// TIA Portal project "Test_PID_Compact_Factory_Cuve" (V16)

(* hardware
DEVICE "Station S7-1200_1"  S7-1200 Station
   slot 0: "Châssis_0"  S7-1200 Rack  Rack  V1.0
   slot 1: "PLC_1"  CPU 1212C DC/DC/DC  6ES7 212-1AE40-0XB0  V4.4
DEVICE "HMI_1"  KTP1200 Basic PN
   slot 0: "HMI_1"  KTP1200 Basic PN  6AV2 123-2MB03-0AX0  16.0.0.0
   slot 1: "HMI_RT_1"  KTP1200 Basic PN  6AV2 123-2MB03-0AX0  16.0.0.0
   slot 5: "HMI_1.IE_CP_1"  PROFINET Interface  16.0.0.0
      slot 1: "Interface PROFINET_1"  PROFINET Interface
         slot 1: "Port_1"  Port
*)

// ===== PLC "PLC_1"  CPU 1212C DC/DC/DC =====

VAR_GLOBAL   // PLC tag table "Table de variables standard"
   "Clock_Byte" AT %MB1000 : Byte;
   "Clock_10Hz" AT %M1000.0 : Bool;
   "Clock_5Hz" AT %M1000.1 : Bool;
   "Clock_2.5Hz" AT %M1000.2 : Bool;
   "Clock_2Hz" AT %M1000.3 : Bool;
   "Clock_1.25Hz" AT %M1000.4 : Bool;
   "Clock_1Hz" AT %M1000.5 : Bool;
   "Clock_0.625Hz" AT %M1000.6 : Bool;
   "Clock_0.5Hz" AT %M1000.7 : Bool;
   "Bouton_0" AT %I0.0 : Bool;
   "Bouton_1" AT %I0.1 : Bool;
   "Bouton_2" AT %I0.2 : Bool;
   "Bouton_3" AT %I0.3 : Bool;
   "Bouton_4" AT %I0.4 : Bool;
   "Bouton_5" AT %I0.5 : Bool;
   "Bouton_6" AT %I0.6 : Bool;
   "Bouton_7" AT %I0.7 : Bool;
   "Sortie_0" AT %Q0.0 : Bool;
   "Sortie_1" AT %Q0.1 : Bool;
   "Sortie_2" AT %Q0.2 : Bool;
   "Sortie_3" AT %Q0.3 : Bool;
   "Sortie_4" AT %Q0.4 : Bool;
   "Sortie_5" AT %Q0.5 : Bool;
   "Commande_Vanne_pcent" AT %MD6 : Real;
   "Consigne_Niveau_Litres" AT %MD10 : Real;
   "Bruit" AT %MD18 : Real;
   "Erreur_Niveau_Litres" AT %MD22 : Real;
   "Correcteur_P_Coeff" AT %MD30 : Real;
   "Erreur_Niveau_pcent" AT %MD26 : Real;
   "Limite_Commande_Max_pcent" AT %MD34 : Real;
   "Limite_Commande_Min_pcent" AT %MD38 : Real;
   "Commande_Max_Atteinte" AT %M70.0 : Bool;
   "Commande_Min_Atteinte" AT %M70.1 : Bool;
   "Consigne_Niveau_Auto_Max" AT %MD42 : Real;
   "Consigne_Niveau_Auto_Min" AT %MD46 : Real;
   "Duree_Demi_Cycle" AT %MD50 : Time;
   "Duree_Demi_Cycle_sec" AT %MW54 : Int;
   "Correcteur_Ti_Valeur_sec" AT %MD72 : Real;
   "Correcteur_Td_Valeur_sec" AT %MD76 : Real;
   "Correcteur_KP_pondere" AT %MD80 : Real;
   "Correcteur_Td_pondere" AT %MD84 : Real;
   "Correcteur_Fo_PB_Derive" AT %MD88 : Real;
   "Commande_Evacuation_pcent" AT %MD14 : Real;
   "Niveau_Litres" AT %MD92 : Real;
   "Debit_Entree_lpars" AT %MD200 : Real;
   "Debit_Sortie_lpars" AT %MD204 : Real;
   "Correcteur_Coeff_Disturbance" AT %MD208 : Real;
END_VAR

VAR_GLOBAL   // PLC tag table "Table de variables IHM"
   "IHM_Bouton_Oscillo_1" AT %M100.0 : Bool;
   "IHM_Bouton_Oscillo_2" AT %M100.1 : Bool;
   "IHM_Bouton_PID_ON_OFF" AT %M100.2 : Bool;
   "IHM_Bouton_Limit_ON_OFF" AT %M100.3 : Bool;
   "IHM_Bouton_Boucle_Fermee" AT %M100.4 : Bool;
   "IHM_Bouton_Bruit" AT %M100.5 : Bool;
   "IHM_Affichage_Oscillo_2" AT %M112.0 : Bool;
   "IHM_Bouton_Marche_Auto" AT %M100.6 : Bool;
   "IHM_Affichage_Correcteur" AT %M112.1 : Bool;
   "IHM_Affichage_Correcteur_I" AT %M112.4 : Bool;
   "IHM_Affichage_Correcteur_D" AT %M112.5 : Bool;
   "IHM_Bouton_Correcteur_I" AT %M112.2 : Bool;
   "IHM_Bouton_Correcteur_D" AT %M112.3 : Bool;
   "IHM_Curseur_Correcteur_I" AT %M112.6 : Bool;
   "IHM_Curseur_Correcteur_D" AT %M112.7 : Bool;
   "IHM_Curseur_Correcteur_P" AT %M113.1 : Bool;
   "IHM_Affichage_Tuyau_Arrivee" AT %M113.2 : Bool;
   "IHM_Affichage_Tuyau_Evacuation" AT %M113.3 : Bool;
   "IHM_Deplacement_Fleche_Tuyau_Arrivee" AT %MW114 : Int;
   "IHM_Deplacement_Fleche_Tuyau_Evacuation" AT %MW116 : Int;
   "IHM_Bouton_Disturbance" AT %M113.4 : Bool;
   "IHM_Affichage_Correcteur_A" AT %M113.5 : Bool;
   "IHM_Valeur_Disturbance" AT %MD120 : Real;
END_VAR

VAR_GLOBAL   // PLC tag table "Table de variables Factory"
   "Niveau_Cuve_Factory" AT %IW100 : Int;
   "Commande_Vanne_Factory" AT %QW100 : Int;
   "Commande_Evacuation_Factory" AT %QW102 : Int;
   "Debit_Sortie_Factory" AT %IW102 : Int;
   "Warning_Light" AT %Q200.0 : Bool;
END_VAR

// folder: Régulateur

DATA_BLOCK "Regulation_DB"   // DB2
{ S7_Optimized_Access := 'TRUE' }
VERSION : 0.1
// stored: InstanceOfName Regulation
"Regulation"
BEGIN
END_DATA_BLOCK

// folder: Simulation Systeme

DATA_BLOCK "POV_DB"   // DB1
{ S7_Optimized_Access := 'TRUE' }
VERSION : 0.1
// stored: InstanceOfName POV
"POV"
BEGIN
END_DATA_BLOCK

// folder: Régulateur

FUNCTION_BLOCK "Regulation"   // FB2, LAD
{ S7_Optimized_Access := 'TRUE' }
VERSION : 0.1
   VAR_TEMP
      Commande_Anticipatrice : Real;
   END_VAR
BEGIN

REGION Network 1 (SCL): Commande Anticipatrice
   IF "IHM_Bouton_Disturbance" THEN
       IF "Erreur_Niveau_Litres">=-1.0 THEN
           #Commande_Anticipatrice := "Debit_Sortie_lpars" * "Correcteur_Coeff_Disturbance";
       ELSE
           #Commande_Anticipatrice := 0;
       END_IF;
   ELSE
       #Commande_Anticipatrice := 0;
   END_IF;

   "IHM_Valeur_Disturbance" := #Commande_Anticipatrice;
END_REGION

REGION Network 2: Bloc fonction PID_Compact
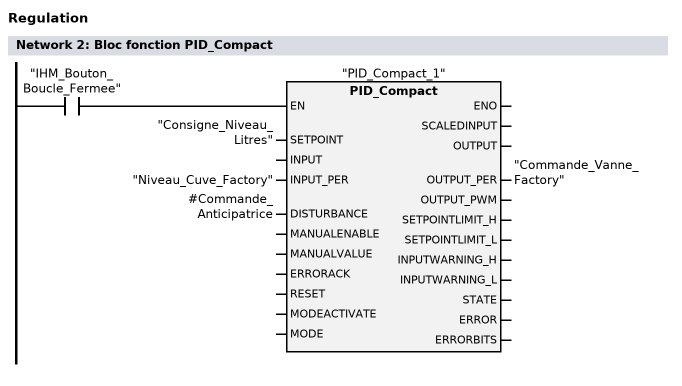
   IF "IHM_Bouton_Boucle_Fermee" THEN
       "PID_Compact_1"(Setpoint := "Consigne_Niveau_Litres",   // PID_Compact
                       Input_PER := "Niveau_Cuve_Factory",
                       Disturbance := #Commande_Anticipatrice,
                       Output_PER => "Commande_Vanne_Factory");
   END_IF;
END_REGION

REGION Network 3 (SCL): Affectation grandeur de commande BO/BF
   // ==== Commande BO / BF ==============================================================================================================
   IF "IHM_Bouton_Boucle_Fermee" THEN
       "Commande_Vanne_pcent":=(INT_TO_REAL("Commande_Vanne_Factory")/27648.0)*100.0;
       "Niveau_Litres" := "PID_Compact_1".ScaledInput;
   ELSE
       "Commande_Vanne_pcent" := "Consigne_Niveau_Litres" ; // Pas des vrais litres...
       "Commande_Vanne_Factory" := REAL_TO_INT("Commande_Vanne_pcent" * 27648.0 / 100.0);
       "Erreur_Niveau_Litres" := 0.0;
       "Erreur_Niveau_pcent" := 0.0;
       "Niveau_Litres" := 300.0 * INT_TO_REAL("Niveau_Cuve_Factory") / 27648.0;
   END_IF;



   // ==== Gestion des limitations de commande ============================================================================================
   REGION Limitations_Commande
       IF "Commande_Vanne_pcent">= "Limite_Commande_Max_pcent" THEN
           "Commande_Vanne_pcent" := "Limite_Commande_Max_pcent";
           "Commande_Max_Atteinte" := "IHM_Bouton_Limit_ON_OFF";
       ELSE
           "Commande_Max_Atteinte" := FALSE;
       END_IF;
       IF "Commande_Vanne_pcent" <= "Limite_Commande_Min_pcent" THEN
           "Commande_Vanne_pcent" := "Limite_Commande_Min_pcent";
           "Commande_Min_Atteinte" := "IHM_Bouton_Limit_ON_OFF";
       ELSE
           "Commande_Min_Atteinte" := FALSE;
       END_IF;
   END_REGION
END_REGION

REGION Network 4 (SCL): Pour affichage IHM
   // ---- Calcul Erreur
   "Erreur_Niveau_Litres" := "Consigne_Niveau_Litres" - "PID_Compact_1".ScaledInput ;
   IF "Consigne_Niveau_Litres" <> 0.0 THEN
       "Erreur_Niveau_pcent" := ("Erreur_Niveau_Litres" / "Consigne_Niveau_Litres") * 100.0;
   ELSE
       "Erreur_Niveau_pcent" := 0.0;
   END_IF;
END_REGION
END_FUNCTION_BLOCK

ORGANIZATION_BLOCK "Appel_Regulation"   // OB32, LAD, CyclicInterrupt
{ S7_Optimized_Access := 'TRUE' }
VERSION : 0.1
   VAR_INPUT
      Initial_Call : Bool;   // Initial call of this OB
      Event_Count : Int;   // Events discarded
   END_VAR
BEGIN

REGION Network 1
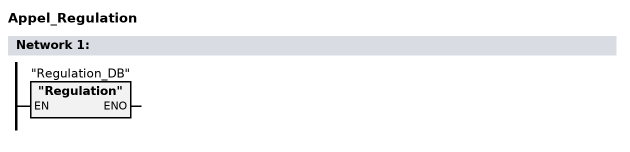
   RUNG wire#powerrail
      "Regulation_DB"()
   END_RUNG
   // the same network as SCL:
   "Regulation_DB"();   // "Regulation"
END_REGION
END_ORGANIZATION_BLOCK

// folder: Simulation Systeme

FUNCTION_BLOCK "POV"   // FB1, LAD
{ S7_Optimized_Access := 'TRUE' }
VERSION : 0.1
   VAR
      Coeff_Perte_Vitesse : Real := 0.3;   // Si 0,4 Perte de 40%
      Temps_Cycle : TON_TIME;
      Temps_Cycle_Demi : TP_TIME;
      Pulse_Cycle : Bool;
   END_VAR
   VAR_TEMP
      Duree_Cycle : Time;
   END_VAR
BEGIN

REGION Network 1 (SCL)
   // ===== Limitations saisie utilisateur IHM =================================================================================

   REGION Limitations_Saisies
       IF "IHM_Bouton_Boucle_Fermee" THEN
           IF "Consigne_Niveau_Litres" > 300.0 THEN
               "Consigne_Niveau_Litres" := 300.0;  // Des vrais litres
           END_IF;
       ELSE
           IF "Consigne_Niveau_Litres" > 100.0 THEN
               "Consigne_Niveau_Litres" := 100.0;  // Pas des litres, mais un pourcentage d'ouverture de la vanne
           END_IF;
           ;
       END_IF;

       IF "Consigne_Niveau_Litres" < 0 THEN
           "Consigne_Niveau_Litres" := 0.0;
       END_IF;

       IF "Commande_Evacuation_pcent" > 100.0 THEN
           "Commande_Evacuation_pcent" := 100.0;
       END_IF;
       IF "Commande_Evacuation_pcent" <0  THEN
           "Commande_Evacuation_pcent" := 0.0;
       END_IF;
   END_REGION


   // ===== Evacuation et débits E/S ===========================================================================================
   "Commande_Evacuation_Factory" := REAL_TO_INT(("Commande_Evacuation_pcent" / 100.0) * 27648.0);
   "Debit_Sortie_lpars":= 9.93*(INT_TO_REAL("Debit_Sortie_Factory")/27648.0);
   "Debit_Entree_lpars" := 7.0 * "Commande_Vanne_pcent" / 100.0;

   // ===== Affichage IHM ======================================================================================================
   REGION Affichage_IHM

       "IHM_Affichage_Oscillo_2" := "IHM_Bouton_Oscillo_2" AND "IHM_Bouton_Oscillo_1";
       "IHM_Affichage_Correcteur" := "IHM_Bouton_Boucle_Fermee" AND "IHM_Bouton_PID_ON_OFF";
       "IHM_Affichage_Correcteur_I" := "IHM_Affichage_Correcteur" AND "IHM_Bouton_Correcteur_I";
       "IHM_Affichage_Correcteur_D" := "IHM_Affichage_Correcteur" AND "IHM_Bouton_Correcteur_D";
       "IHM_Affichage_Correcteur_A" := "IHM_Affichage_Correcteur" AND "IHM_Bouton_Disturbance";

       IF (("Correcteur_Ti_Valeur_sec" <> 0) AND "IHM_Affichage_Correcteur_I" ) THEN
           "IHM_Curseur_Correcteur_I" := TRUE;
       ELSE
           "IHM_Curseur_Correcteur_I" := FALSE;
       END_IF;
       IF (("Correcteur_Td_Valeur_sec" <> 0) AND "IHM_Affichage_Correcteur_D" ) THEN
           "IHM_Curseur_Correcteur_D" := TRUE;
       ELSE
           "IHM_Curseur_Correcteur_D" := FALSE;
       END_IF;

       IF "IHM_Affichage_Correcteur" THEN
           "IHM_Curseur_Correcteur_P" := TRUE;
       ELSE
           "IHM_Curseur_Correcteur_P" := FALSE;
       END_IF;

       "Correcteur_P_Coeff" := "PID_Compact_1".#Retain.CtrlParams.Gain ;
       "Correcteur_KP_pondere" := "PID_Compact_1".#Retain.CtrlParams.Gain * "PID_Compact_1".Retain.CtrlParams.PWeighting;
       "Correcteur_Ti_Valeur_sec" := "PID_Compact_1".Retain.CtrlParams.Ti;
       "Correcteur_Td_Valeur_sec" := "PID_Compact_1".Retain.CtrlParams.Td;
       "Correcteur_Td_pondere" := "PID_Compact_1".Retain.CtrlParams.Td * "PID_Compact_1".Retain.CtrlParams.DWeighting;
       "Correcteur_Fo_PB_Derive" := 1.0 / (2 * 3.1415927 * "PID_Compact_1".Retain.CtrlParams.TdFiltRatio * "Correcteur_Td_Valeur_sec");

       IF "Commande_Vanne_pcent" > 0.0 THEN
           "IHM_Affichage_Tuyau_Arrivee" := TRUE;
       ELSE
           "IHM_Affichage_Tuyau_Arrivee" := FALSE;
       END_IF;
       IF "Debit_Sortie_lpars" > 0.1 THEN
           "IHM_Affichage_Tuyau_Evacuation" := TRUE;
       ELSE
           "IHM_Affichage_Tuyau_Evacuation" := FALSE;
       END_IF;

       IF "Niveau_Litres">280.0 THEN
           "Warning_Light" := TRUE;
       ELSE
           "Warning_Light" := FALSE;
       END_IF;



   END_REGION



   // ===== Marche AUTO consigne créneau =======================================================================================
   REGION Creneau_Consigne
       IF "IHM_Bouton_Marche_Auto" THEN
           IF NOT #Temps_Cycle_Demi.Q THEN
               "Consigne_Niveau_Litres" := "Consigne_Niveau_Auto_Max";
           END_IF;
           IF #Temps_Cycle_Demi.Q THEN
               "Consigne_Niveau_Litres" := "Consigne_Niveau_Auto_Min";
           END_IF;
       END_IF;
       "Duree_Demi_Cycle" := INT_TO_TIME("Duree_Demi_Cycle_sec" * 1000);
       #Duree_Cycle := "Duree_Demi_Cycle" * 2;
   END_REGION
END_REGION

REGION Network 2: Tempo Cycle Auto
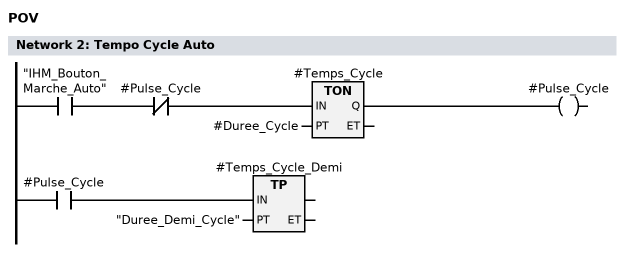
   #Temps_Cycle(IN := "IHM_Bouton_Marche_Auto" AND NOT #Pulse_Cycle, PT := #Duree_Cycle);   // TON
   #Pulse_Cycle := #Temps_Cycle.Q;
   #Temps_Cycle_Demi(IN := #Pulse_Cycle, PT := "Duree_Demi_Cycle");   // TP
END_REGION
END_FUNCTION_BLOCK

ORGANIZATION_BLOCK "Main"   // OB1, LAD, ProgramCycle
TITLE = "Main Program Sweep (Cycle)"
{ S7_Optimized_Access := 'TRUE' }
VERSION : 0.1
   VAR_INPUT
      Initial_Call : Bool;   // Initial call of this OB
      Remanence : Bool;   // =True, if remanent data are available
   END_VAR
BEGIN

REGION Network 1: Appel fonction de simulation de la partie opérative
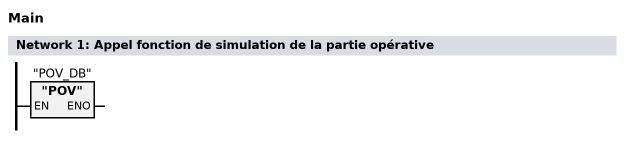
   RUNG wire#powerrail
      "POV_DB"()
   END_RUNG
   // the same network as SCL:
   "POV_DB"();   // "POV"
END_REGION
END_ORGANIZATION_BLOCK

ORGANIZATION_BLOCK "Affichage_Fleches"   // OB30, LAD, CyclicInterrupt
{ S7_Optimized_Access := 'TRUE' }
VERSION : 0.1
   VAR_INPUT
      Initial_Call : Bool;   // Initial call of this OB
      Event_Count : Int;   // Events discarded
   END_VAR
   VAR_TEMP
      Increment_Arrivee : Int;
      Increment_Evacuation : Int;
   END_VAR
BEGIN

REGION Network 1 (SCL)
   #Increment_Arrivee := REAL_TO_INT("Commande_Vanne_pcent" / 5.0) ;
   "IHM_Deplacement_Fleche_Tuyau_Arrivee" := "IHM_Deplacement_Fleche_Tuyau_Arrivee" + #Increment_Arrivee;
   IF "IHM_Deplacement_Fleche_Tuyau_Arrivee" > 100 THEN
       "IHM_Deplacement_Fleche_Tuyau_Arrivee" := 0;
   END_IF;

   #Increment_Evacuation := REAL_TO_INT("Debit_Sortie_lpars" * 2.0);
   "IHM_Deplacement_Fleche_Tuyau_Evacuation" := "IHM_Deplacement_Fleche_Tuyau_Evacuation" + #Increment_Evacuation;
   IF "IHM_Deplacement_Fleche_Tuyau_Evacuation" > 100 THEN
       "IHM_Deplacement_Fleche_Tuyau_Evacuation" := 0;
   END_IF;
END_REGION
END_ORGANIZATION_BLOCK

ORGANIZATION_BLOCK "Startup"   // OB100, LAD, Startup
TITLE = "Complete Restart"
{ S7_Optimized_Access := 'TRUE' }
VERSION : 0.1
   VAR_INPUT
      LostRetentive : Bool;   // True if retentive data are lost
      LostRTC : Bool;   // True if date and time are lost
   END_VAR
BEGIN

REGION Network 1 (SCL): Valeurs Initiales du système et du régulateur

   "Limite_Commande_Max_pcent" := 100.0;
   "Limite_Commande_Min_pcent" := 0.0;

   "Consigne_Niveau_Auto_Max" := 200.0;
   "Consigne_Niveau_Auto_Min" := 100.0;

   "Duree_Demi_Cycle_sec" := 5;

   "Correcteur_Coeff_Disturbance" := 1;
END_REGION
END_ORGANIZATION_BLOCK

(* ===== HMI "HMI_RT_1" =====
system functions are stored by id; their names below are inferred from use
connection "HMI_Liaison_1": ETHERNET, SMART_S7_1200_OMS

HMI tags "Table de variables standard"
   "IHM_Bouton_Oscillo_2" : Bool = PLC IHM_Bouton_Oscillo_2 AT %M100.1, 500 ms
   "IHM_Bouton_PID_ON_OFF" : Bool = PLC IHM_Bouton_PID_ON_OFF AT %M100.2, 500 ms
   "IHM_Bouton_Boucle_Fermee" : Bool = PLC IHM_Bouton_Boucle_Fermee AT %M100.4, 500 ms
   "Niveau_Litres" : Real = PLC Niveau_Litres AT %MD92, 100 ms
   "Evacuation_pcent" : Real = PLC Commande_Evacuation_pcent AT %MD14, 100 ms
   "Commande_Vanne_pcent" : Real = PLC Commande_Vanne_pcent AT %MD6, 100 ms
   "IHM_Bouton_Oscillo_1" : Bool = PLC IHM_Bouton_Oscillo_1 AT %M100.0, 500 ms
   "Consigne_Niveau_Litres" : Real = PLC Consigne_Niveau_Litres AT %MD10, 100 ms
   "IHM_Bouton_Bruit" : Bool = PLC IHM_Bouton_Bruit AT %M100.5, 500 ms
   "Erreur_Niveau_Litres" : Real = PLC Erreur_Niveau_Litres AT %MD22, 100 ms
   "Erreur_Niveau_pcent" : Real = PLC Erreur_Niveau_pcent AT %MD26, 100 ms
   "Correcteur_P_Coeff" : Real = PLC Correcteur_P_Coeff AT %MD30, 500 ms
   "IHM_Bouton_Limit_ON_OFF" : Bool = PLC IHM_Bouton_Limit_ON_OFF AT %M100.3, 500 ms
   "Limite_Commande_Max_pcent" : Real = PLC Limite_Commande_Max_pcent AT %MD34, 1 s
   "Limite_Commande_Min_pcent" : Real = PLC Limite_Commande_Min_pcent AT %MD38, 1 s
   "Commande_Max_Atteinte" : Bool = PLC Commande_Max_Atteinte AT %M70.0, 100 ms
   "Commande_Min_Atteinte" : Bool = PLC Commande_Min_Atteinte AT %M70.1, 100 ms
   "IHM_Affichage_Oscillo_2" : Bool = PLC IHM_Affichage_Oscillo_2 AT %M112.0, 500 ms
   "IHM_Bouton_Marche_Auto" : Bool = PLC IHM_Bouton_Marche_Auto AT %M100.6, 500 ms
   "Consigne_Niveau_Auto_Max" : Real = PLC Consigne_Niveau_Auto_Max AT %MD42, 1 s
   "Consigne_Niveau_Auto_Min" : Real = PLC Consigne_Niveau_Auto_Min AT %MD46, 1 s
   "Duree_Demi_Cycle_sec" : Int = PLC Duree_Demi_Cycle_sec AT %MW54, 1 s
   "OV_DB.Temps_Cycle.ET" : Time = PLC POV_DB.Temps_Cycle.ET, 100 ms
   "IHM_Affichage_Correcteur" : Bool = PLC IHM_Affichage_Correcteur AT %M112.1, 500 ms
   "Correcteur_Ti_Valeur_sec" : Real = PLC Correcteur_Ti_Valeur_sec AT %MD72, 500 ms
   "Correcteur_Td_Valeur_sec" : Real = PLC Correcteur_Td_Valeur_sec AT %MD76, 500 ms
   "IHM_Bouton_Correcteur_I" : Bool = PLC IHM_Bouton_Correcteur_I AT %M112.2, 1 s
   "IHM_Bouton_Correcteur_D" : Bool = PLC IHM_Bouton_Correcteur_D AT %M112.3, 1 s
   "IHM_Affichage_Correcteur_D" : Bool = PLC IHM_Affichage_Correcteur_D AT %M112.5, 500 ms
   "IHM_Affichage_Correcteur_I" : Bool = PLC IHM_Affichage_Correcteur_I AT %M112.4, 500 ms
   "IHM_Bouton_Oscillo_Erreur" : Bool AT %DB1.DBX0.0
   "IHM_Curseur_Correcteur_I" : Bool = PLC IHM_Curseur_Correcteur_I AT %M112.6, 500 ms
   "IHM_Curseur_Correcteur_D" : Bool = PLC IHM_Curseur_Correcteur_D AT %M112.7, 500 ms
   "IHM_Curseur_Correcteur_P" : Bool = PLC IHM_Curseur_Correcteur_P AT %M113.1, 500 ms
   "Correcteur_Td_pondere" : Real = PLC Correcteur_Td_pondere AT %MD84, 500 ms
   "Correcteur_KP_pondere" : Real = PLC Correcteur_KP_pondere AT %MD80, 500 ms
   "Correcteur_Fo_PB_Derive" : Real = PLC Correcteur_Fo_PB_Derive AT %MD88, 500 ms
   "IHM_Affichage_Tuyau_Evacuation" : Bool = PLC IHM_Affichage_Tuyau_Evacuation AT %M113.3, 100 ms
   "IHM_Affichage_Tuyau_Arrivee" : Bool = PLC IHM_Affichage_Tuyau_Arrivee AT %M113.2, 100 ms
   "Debit_Sortie_lpars" : Real = PLC Debit_Sortie_lpars AT %MD204, 100 ms
   "Bouton_Affichage_Debit_Sortie" : Bool AT %DB1.DBD0
   "Bouton_Affichage_Debit_Entree" : Bool AT %DB1.DBD0
   "Debit_Entree_lpars" : Real = PLC Debit_Entree_lpars AT %MD200, 100 ms
   "IHM_Deplacement_Fleche_Tuyau_Arrivee" : Int = PLC IHM_Deplacement_Fleche_Tuyau_Arrivee AT %MW114, 100 ms
   "IHM_Deplacement_Fleche_Tuyau_Evacuation" : Int = PLC IHM_Deplacement_Fleche_Tuyau_Evacuation AT %MW116, 100 ms
   "IHM_Bouton_Disturbance" : Bool = PLC IHM_Bouton_Disturbance AT %M113.4, 500 ms
   "Correcteur_Coeff_Disturbance" : Real = PLC Correcteur_Coeff_Disturbance AT %MD208, 500 ms
   "IHM_Affichage_Correcteur_A" : Bool = PLC IHM_Affichage_Correcteur_A AT %M113.5, 500 ms
   "IHM_Valeur_Disturbance" : Real = PLC IHM_Valeur_Disturbance AT %MD120, 100 ms

text list "Liste de textes_1": 1 'Ordre 1'; 2 'Ordre 2'; 3 'Ordre 2+1'

text list "Liste de textes_Correcteur_Mixte": 0 'Parallèle'; 1 'Mixte'

screen "Vue racine" 1280x800, template "Modèle_1"
   TextField "HmiScreenItemData_1" at 236,261 size 12x25; Text '-'
   TextField "HmiScreenItemData_14" at 218,244 size 19x25; Text '+'
   TextField "HmiScreenItemData_16" at 133,342 size 63x25; Text 'Boucle'
   TextField "HmiScreenItemData_15" at 131,370 size 68x25; Text 'Fermée'
   GraphicView "Vue de graphique_27" at 911,0 size 33x61; Picture "Graphique_89"
   GraphicView "Vue de graphique_7" at 942,34 size 52x52; Picture "Graphique_180"
   GraphicView "Vue de graphique_22" at 1087,349 size 68x68; Picture "Graphique_174"
   GraphicView "Vue de graphique_2" at 1148,349 size 132x68; Picture "Graphique_166"
   GraphicView "Vue de graphique_4" at 939,47 size 226x353; Picture "Graphique_125"
   Rectangle "Rectangle_2" at 412,189 size 168x211
      Visibility <- "IHM_Affichage_Correcteur"
   Line "Ligne_5" at 242,500 size 807x0
      Visibility <- "IHM_Bouton_Boucle_Fermee"
   GraphicView "Vue de graphique_15" at 225,273 size 36x30; Picture "Graphique_106"
      Visibility <- "IHM_Bouton_Boucle_Fermee"
   Line "Ligne_1" at 1051,381 size 0x119
      Visibility <- "IHM_Bouton_Boucle_Fermee"
   GraphicView "Vue de graphique_14" at 194,244 size 36x30; Picture "Graphique_104"
   TextField "HmiScreenItemData_7" at 1083,412 size 80x27; Text 'Litres'
   GraphicView "Vue de graphique_11" at 702,140 size 27x27; Picture "Graphique_60"
      Visibility <- "Commande_Max_Atteinte"
   TrendView "Vue de courbes_1" at 660,457 size 620x343
      Visibility <- "IHM_Bouton_Oscillo_1"
   Button "Bouton_5" at 1037,373 size 28x15; TextOff 'Text'; PictureOff "Graphique_98"
      on Click: InvertBit("IHM_Bouton_Oscillo_1")
   GraphicView "Vue de graphique_13" at 767,244 size 36x30; Picture "Graphique_104"
   TextField "HmiScreenItemData_6" at 1013,354 size 76x17; Text 'Mesure Niveau'
   IOField "Champ d'E/S_2" at 1002,409 size 97x32; FormatPattern 999.9
      ProcessValue <- "Niveau_Litres"
   Group "Group_4" at 216,231 size 53x55
   Group "Group_5" at 131,342 size 68x53
   Line "Ligne_6" at 242,283 size 0x217
      Visibility <- "IHM_Bouton_Boucle_Fermee"
   Switch "Commutateur_1" at 212,355 size 64x32; CaptionText 'Switch'; TextOff 'OFF'; TextOn 'ON'
      ProcessValue <- "IHM_Bouton_Boucle_Fermee"
   Rectangle "Rectangle_1" at 194,218 size 97x91
      Visibility <- "IHM_Bouton_Boucle_Fermee"
   Line "Ligne_7" at 193,258 size 103x0
      Visibility <- "IHM_Bouton_Boucle_Fermee"
   TextField "HmiScreenItemData_17" at 297,228 size 53x22; Text 'Erreur'
      Visibility <- "IHM_Bouton_Boucle_Fermee"
   IOField "Champ d'E/S_3" at 288,270 size 71x22; FormatPattern s999.9
      ProcessValue <- "Erreur_Niveau_Litres"
      Visibility <- "IHM_Bouton_Boucle_Fermee"
   IOField "Champ d'E/S_6" at 288,300 size 71x22; FormatPattern s999.99
      ProcessValue <- "Erreur_Niveau_pcent"
      Visibility <- "IHM_Bouton_Boucle_Fermee"
   TextField "HmiScreenItemData_18" at 360,271 size 34x18; Text 'Litres'
      Visibility <- "IHM_Bouton_Boucle_Fermee"
   TextField "HmiScreenItemData_19" at 361,301 size 17x18; Text '%'
      Visibility <- "IHM_Bouton_Boucle_Fermee"
   IOField "Champ d'E/S_7" at 454,201 size 71x22; FormatPattern 999.9
      ProcessValue <- "Correcteur_P_Coeff"
      Visibility <- "IHM_Affichage_Correcteur"
   Button "Bouton_7" at 707,253 size 18x11; TextOff 'Text'; PictureOff "Graphique_98"
      on Click: InvertBit("IHM_Bouton_Limit_ON_OFF")
   Line "Ligne_8" at 716,209 size 0x41
      Visibility <- "IHM_Bouton_Limit_ON_OFF"
   Line "Ligne_9" at 710,208 size 12x0
      Visibility <- "IHM_Bouton_Limit_ON_OFF"
   Line "Ligne_10" at 716,267 size 0x41
      Visibility <- "IHM_Bouton_Limit_ON_OFF"
   Line "Ligne_11" at 710,308 size 12x0
      Visibility <- "IHM_Bouton_Limit_ON_OFF"
   IOField "Champ d'E/S_8" at 680,182 size 71x22; FormatPattern s9999
      ProcessValue <- "Limite_Commande_Max_pcent"
      Visibility <- "IHM_Bouton_Limit_ON_OFF"
   IOField "Champ d'E/S_9" at 680,314 size 71x22; FormatPattern s9999
      ProcessValue <- "Limite_Commande_Min_pcent"
      Visibility <- "IHM_Bouton_Limit_ON_OFF"
   GraphicView "Vue de graphique_16" at 702,350 size 27x27; Picture "Graphique_60"
      Visibility <- "Commande_Min_Atteinte"
   Button "Bouton_8" at 479,252 size 18x11; TextOff 'Text'; PictureOff "Graphique_98"
      on Click: InvertBit("IHM_Bouton_PID_ON_OFF")
      Visibility <- "IHM_Bouton_Boucle_Fermee"
   TextField "HmiScreenItemData_20" at 424,210 size 15x22; Text 'P'
      Visibility <- "IHM_Affichage_Correcteur"
   TextField "HmiScreenItemData_21" at 458,164 size 86x22; Text 'Correcteur'
      Visibility <- "IHM_Affichage_Correcteur"
   IOField "Champ d'E/S_5" at 24,243 size 96x32; FormatPattern 999
      ProcessValue <- "Consigne_Niveau_Litres"
   Button "Bouton_9" at 138,229 size 22x22; TextOff '+'
      on Press: function_dd21b452("Consigne_Niveau_Litres", 20)
   Bar "Bargraphe_1" at 48,32 size 54x200; MinimumValue 0; MaximumValue 300
      ProcessValue <- "Consigne_Niveau_Litres"
      Visibility <- "IHM_Bouton_Boucle_Fermee"
   Button "Bouton_10" at 138,266 size 22x22; TextOff '-'
      on Press: function_dd21b452("Consigne_Niveau_Litres", -20)
   Button "Bouton_11" at 621,742 size 35x32; TextOff 'Text'; PictureOff "Graphique_114"
      on Click: InvertBit("IHM_Bouton_Oscillo_2")
      Visibility <- "IHM_Bouton_Oscillo_1"
   Switch "Commutateur_2" at 200,109 size 32x64; CaptionText 'Switch'; TextOff '-'; TextOn '~'
      ProcessValue <- "IHM_Bouton_Marche_Auto"
   TextField "HmiScreenItemData_22" at 272,32 size 33x22; Text 'Max'
      Visibility <- "IHM_Bouton_Marche_Auto"
   IOField "Champ d'E/S_10" at 337,31 size 71x22; FormatPattern 999
      Visibility <- "IHM_Bouton_Marche_Auto"
      ProcessValue <- "Consigne_Niveau_Auto_Max"
   IOField "Champ d'E/S_11" at 337,65 size 71x22; FormatPattern 999
      Visibility <- "IHM_Bouton_Marche_Auto"
      ProcessValue <- "Consigne_Niveau_Auto_Min"
   IOField "Champ d'E/S_12" at 337,100 size 71x22; FormatPattern 999
      Visibility <- "IHM_Bouton_Marche_Auto"
      ProcessValue <- "Duree_Demi_Cycle_sec"
   TextField "HmiScreenItemData_23" at 272,65 size 27x22; Text 'Min'
      Visibility <- "IHM_Bouton_Marche_Auto"
   TextField "HmiScreenItemData_24" at 272,99 size 58x22; Text 'Durée/2'
      Visibility <- "IHM_Bouton_Marche_Auto"
   TextField "HmiScreenItemData_25" at 138,146 size 40x22; Text 'FIXE'
      Visibility <- "IHM_Bouton_Marche_Auto"
   TextField "HmiScreenItemData_26" at 138,111 size 54x22; Text 'CYCLE'
      Visibility <- "IHM_Bouton_Marche_Auto"
   IOField "Champ d'E/S_13" at 454,282 size 71x22; FormatPattern 99999.99
      ProcessValue <- "Correcteur_Ti_Valeur_sec"
      Visibility <- "IHM_Affichage_Correcteur_I"
   TextField "HmiScreenItemData_27" at 424,282 size 12x22; Text 'I'
      Visibility <- "IHM_Affichage_Correcteur_I"
   IOField "Champ d'E/S_14" at 454,324 size 71x22; FormatPattern 9999.999
      ProcessValue <- "Correcteur_Td_Valeur_sec"
      Visibility <- "IHM_Affichage_Correcteur_D"
   TextField "HmiScreenItemData_28" at 423,334 size 16x22; Text 'D'
      Visibility <- "IHM_Affichage_Correcteur_D"
   TextField "HmiScreenItemData_29" at 527,286 size 17x14; Text 'sec'
      Visibility <- "IHM_Affichage_Correcteur_I"
   TextField "HmiScreenItemData_30" at 526,328 size 28x14; Text 'Retour'
      Visibility <- "IHM_Affichage_Correcteur_D"
   TextField "HmiScreenItemData_31" at 688,164 size 55x17; Text 'Limite Max'
      Visibility <- "IHM_Bouton_Limit_ON_OFF"
   TextField "HmiScreenItemData_32" at 690,335 size 51x17; Text 'Limite Min'
      Visibility <- "IHM_Bouton_Limit_ON_OFF"
   Rectangle "Rectangle_3" at 51,737 size 561x19
      Visibility <- "IHM_Affichage_Oscillo_2"
   IOField "Champ d'E/S_17" at 422,100 size 55x22; FormatPattern 999999
      Visibility <- "IHM_Bouton_Marche_Auto"
      ProcessValue <- "OV_DB.Temps_Cycle.ET"
   TextField "HmiScreenItemData_35" at 453,100 size 24x22; Text 'Sec'
      Visibility <- "IHM_Bouton_Marche_Auto"
   Button "Bouton_17" at 138,294 size 22x11; TextOff '0'; PictureOff "Graphique_98"
      on Click: SetTag("Consigne_Niveau_Litres", 0)
   Button "Bouton_18" at 138,212 size 22x11; TextOff '200'; PictureOff "Graphique_98"
      on Click: SetTag("Consigne_Niveau_Litres", 200)
      Visibility <- "IHM_Bouton_Boucle_Fermee"
   Button "Bouton_19" at 408,286 size 10x16; TextOff 'Text'; PictureOff "Graphique_98"
      on Click: InvertBit("IHM_Bouton_Correcteur_I")
      Visibility <- "IHM_Affichage_Correcteur"
   Button "Bouton_20" at 408,337 size 10x16; TextOff 'Text'; PictureOff "Graphique_98"
      on Click: InvertBit("IHM_Bouton_Correcteur_D")
      Visibility <- "IHM_Affichage_Correcteur"
   Button "Bouton_21" at 316,253 size 18x11; TextOff 'Text'; PictureOff "Graphique_98"
      on Click: InvertBit("IHM_Bouton_Oscillo_Erreur")
      Visibility <- "IHM_Bouton_Boucle_Fermee"
   IOField "Champ d'E/S_19" at 454,225 size 71x22; FormatPattern 999.9
      Visibility <- "IHM_Affichage_Correcteur"
      ProcessValue <- "Correcteur_KP_pondere"
   TextField "HmiScreenItemData_37" at 525,230 size 36x14; Text 'Consigne'
      Visibility <- "IHM_Affichage_Correcteur"
   TextField "HmiScreenItemData_38" at 526,353 size 36x14; Text 'Consigne'
      Visibility <- "IHM_Affichage_Correcteur_D"
   IOField "Champ d'E/S_20" at 454,348 size 71x22; FormatPattern 9999.999
      Visibility <- "IHM_Affichage_Correcteur_D"
      ProcessValue <- "Correcteur_Td_pondere"
   TextField "HmiScreenItemData_39" at 525,205 size 28x14; Text 'Retour'
      Visibility <- "IHM_Affichage_Correcteur"
   TextField "HmiScreenItemData_5" at 46,321 size 53x25; Text 'Litres'
      Visibility <- "IHM_Bouton_Boucle_Fermee"
   TextField "HmiScreenItemData" at 40,299 size 64x25; Text 'Niveau'
      Visibility <- "IHM_Bouton_Boucle_Fermee"
   TextField "HmiScreenItemData_4" at 30,277 size 84x25; Text 'Consigne'
   TrendView "Vue de courbes_2" at 0,399 size 615x401
      Visibility <- "IHM_Affichage_Oscillo_2"
   TrendView "Vue de courbes_3" at 0,399 size 615x398
      Visibility <- "IHM_Bouton_Oscillo_Erreur"
   GraphicView "Vue de graphique_25" at 1170,358 size 86x50; Picture "Graphique_171"
   GraphicView "Vue de graphique_1" at 859,34 size 52x52; Picture "Graphique_179"
   GraphicView "Vue de graphique_9" at 859,83 size 52x257; Picture "Graphique_185"
   GraphicView "Vue de graphique_8" at 789,237 size 84x48; Picture "Graphique_187"
   GraphicView "Vue de graphique_10" at 867,229 size 36x57; Picture "Graphique_186"
   GraphicView "Vue de graphique_3" at 910,34 size 34x52; Picture "Graphique_166"
   TextField "HmiScreenItemData_13" at 773,134 size 86x22; Text 'Commande'
   TextField "HmiScreenItemData_12" at 791,153 size 51x22; Text 'Vanne'
   TextField "HmiScreenItemData_2" at 768,173 size 97x22; Text 'Arrivée (%)'
   IOField "Champ d'E/S_1" at 772,200 size 88x32; FormatPattern 999.9
      ProcessValue <- "Commande_Vanne_pcent"
   Bar "Bargraphe_2" at 1023,133 size 58x174; MinimumValue 0; MaximumValue 300
      ProcessValue <- "Niveau_Litres"
   GraphicView "Vue de graphique_24" at 789,237 size 84x48; Picture "Graphique_193"
      Visibility <- "IHM_Affichage_Tuyau_Arrivee"
   GraphicView "Vue de graphique_26" at 1247,397 size 33x61; Picture "Graphique_89"
   TextField "HmiScreenItemData_9" at 43,298 size 58x25; Text 'Vanne'
      Visibility <- "IHM_Bouton_Boucle_Fermee"
   TextField "HmiScreenItemData_10" at 60,322 size 25x25; Text '%'
      Visibility <- "IHM_Bouton_Boucle_Fermee"
   Button "Bouton_1" at 138,212 size 22x11; TextOff '100'; PictureOff "Graphique_98"
      on Click: SetTag("Consigne_Niveau_Litres", 100)
      Visibility <- "IHM_Bouton_Boucle_Fermee"
   TextField "HmiScreenItemData_11" at 1184,431 size 70x27; Text 'Litres/sec'
      Visibility <- "Bouton_Affichage_Debit_Sortie"
   Button "Bouton_2" at 1253,419 size 21x10; TextOff 'Text'; PictureOff "Graphique_98"
      on Click: InvertBit("Bouton_Affichage_Debit_Sortie")
   IOField "Champ d'E/S_16" at 947,15 size 53x22; FormatPattern 99.99
      Visibility <- "Bouton_Affichage_Debit_Entree"
      ProcessValue <- "Debit_Entree_lpars"
   TextField "HmiScreenItemData_33" at 991,12 size 70x27; Text 'Litres/sec'
      Visibility <- "Bouton_Affichage_Debit_Entree"
   Button "Bouton_6" at 917,22 size 21x10; TextOff 'Text'; PictureOff "Graphique_98"
      on Click: InvertBit("Bouton_Affichage_Debit_Entree")
   GraphicView "Vue de graphique_30" at 920,40 size 18x41; Picture "Graphique_199"
   GraphicView "Vue de graphique_28" at 1256,354 size 20x54; Picture "Graphique_199"
   GraphicView "Vue de graphique_6" at 840,330 size 90x113; Picture "Graphique_177"
   GraphicView "Vue de graphique_18" at 1133,360 size 44x44; Picture "Graphique_200"
      Visibility <- "IHM_Affichage_Tuyau_Evacuation"
      HorizontalMovement <- "IHM_Deplacement_Fleche_Tuyau_Evacuation"
   IOField "Champ d'E/S_4" at 1177,294 size 71x22; FormatPattern s999.9
      ProcessValue <- "Evacuation_pcent"
   Button "Bouton_4" at 1177,326 size 27x24; TextOff '-'
      on Press: function_dd21b452("Evacuation_pcent", -10)
   Button "Bouton_3" at 1221,326 size 27x24; TextOff '+'
      on Press: function_dd21b452("Evacuation_pcent", 10)
   TextField "HmiScreenItemData_3" at 1163,267 size 99x27; Text 'Evacuation'
   TextField "HmiScreenItemData_8" at 1241,291 size 32x27; Text '%'
   GraphicView "Vue de graphique_5" at 863,167 size 43x43; Picture "Graphique_201"
      Visibility <- "IHM_Affichage_Tuyau_Arrivee"
      VerticalMovement <- "IHM_Deplacement_Fleche_Tuyau_Arrivee"
   GraphicView "Vue de graphique_12" at 863,296 size 43x43; Picture "Graphique_201"
      Visibility <- "IHM_Affichage_Tuyau_Arrivee"
      VerticalMovement <- "IHM_Deplacement_Fleche_Tuyau_Arrivee"
   Button "Bouton_12" at 574,374 size 10x16; TextOff 'Text'; PictureOff "Graphique_98"
      on Click: InvertBit("IHM_Bouton_Disturbance")
      Visibility <- "IHM_Affichage_Correcteur"
   TextField "HmiScreenItemData_34" at 554,370 size 15x22; Text 'A'
      Visibility <- "IHM_Affichage_Correcteur_A"
   Button "Bouton_13" at 588,372 size 17x11; TextOff '+'; PictureOff "Graphique_98"
      on Click: function_dd21b452("Correcteur_Coeff_Disturbance", 1)
      Visibility <- "IHM_Affichage_Correcteur_A"
   Button "Bouton_14" at 588,383 size 17x11; TextOff '-'; PictureOff "Graphique_98"
      on Click: function_dd21b452("Correcteur_Coeff_Disturbance", -1)
      Visibility <- "IHM_Affichage_Correcteur_A"
   Line "Ligne_20" at 643,450 size 535x0
      Visibility <- "IHM_Affichage_Correcteur_A"
   Line "Ligne_21" at 1178,434 size 16x16
      Visibility <- "IHM_Affichage_Correcteur_A"
   IOField "Champ d'E/S_15" at 1191,415 size 55x22; FormatPattern 99.99
      ProcessValue <- "Debit_Sortie_lpars"
      Visibility <- "Bouton_Affichage_Debit_Sortie"
   Group "Group" at 590,212 size 103x87
   Line "Ligne_19" at 642,285 size 0x165
      Visibility <- "IHM_Affichage_Correcteur_A"
   IOField "Champ d'E/S_18" at 608,372 size 71x22
      ProcessValue <- "Correcteur_Coeff_Disturbance"
      Visibility <- "IHM_Affichage_Correcteur_A"
   IOField "Champ d'E/S_21" at 587,295 size 50x22; FormatPattern 999.9
      Visibility <- "IHM_Affichage_Correcteur_A"
      ProcessValue <- "IHM_Valeur_Disturbance"
   TextField "HmiScreenItemData_41" at 586,314 size 53x15; Text 'Disturbance'
      Visibility <- "IHM_Affichage_Correcteur_A"
   TextField "HmiScreenItemData_42" at 645,297 size 17x18; Text '%'
      Visibility <- "IHM_Affichage_Correcteur_A"
   Rectangle "Rectangle_6" at 606,212 size 76x87
      Visibility <- "IHM_Affichage_Correcteur_A"
   Line "Ligne_14" at 590,258 size 103x0
      Visibility <- "IHM_Affichage_Correcteur_A"
   Circle "Cercle_2" at 616,231 size 53x53
      Visibility <- "IHM_Affichage_Correcteur_A"
   Line "Ligne_12" at 625,240 size 35x35
      Visibility <- "IHM_Affichage_Correcteur_A"
   Line "Ligne_13" at 625,240 size 34x34
      Visibility <- "IHM_Affichage_Correcteur_A"
   TextField "HmiScreenItemData_36" at 633,260 size 19x25; Text '+'
      Visibility <- "IHM_Affichage_Correcteur_A"
   TextField "HmiScreenItemData_40" at 618,244 size 19x25; Text '+'
      Visibility <- "IHM_Affichage_Correcteur_A"
   Line "Ligne_15" at 608,252 size 7x5
      Visibility <- "IHM_Affichage_Correcteur_A"
   Line "Ligne_16" at 608,258 size 7x5
      Visibility <- "IHM_Affichage_Correcteur_A"
   Line "Ligne_17" at 643,284 size 5x7
      Visibility <- "IHM_Affichage_Correcteur_A"
   Line "Ligne_18" at 636,284 size 5x7
      Visibility <- "IHM_Affichage_Correcteur_A"
*)